(* IEC 61131-3 sources: SortJet_MasterSPS_Aufbau.fbsproj/Device.device.xml.v3^/Plc Logic.plclogic.xml.v3^/Application.application.xml.v3^/09_Station/Stationen/Förderer[202,203]/0_Konfig, 6 files *)

(* ---- Antriebsinformationen_202.gvl ---- *)
(* METADATA
{
	"v3Meta": {
		"objectGuid": "ae52444f-d7c0-4b01-95e4-d9e00420f7a3"
	}
}
*)
{attribute 'allow_unqualified_access'}
NAMESPACE Antriebsinformationen_202
VAR_GLOBAL

//**************************************************************************************************)
// ANTRIEBSINFORMATION  *)
//**************************************************************************************************)

  apgInfoStation202Glastransport : ARRAY[cWAND_1..cANZAHL_WAENDE] OF AntriebsInformationen := [
    (
      wAchsID                                 :=      12,  // Achs ID aus dem EConSet
      stTyp                                   := 'Belt',  // Typ
      wpSchaltschrank                         :=   2020,  // Daten aus dem Schaltplan
      wpSchaltplanreihe                       :=      2,  // Daten aus dem Schaltplan
      wpSchaltplanseite                       :=    100,  // Daten aus dem Schaltplan
      rpMaxGeschwindigkeit                    :=   1000,  // [mm/s]   Max- Geschwindigkeit für den Automatikbetrieb
      rpHandGeschwindigkeit                   :=    333,  // [mm/s]   Hand- Geschwindigkeit
      rpReduzierteGeschwindigkeit             :=    250,  // [mm/s]   Reduzierte Geschwindigkeit
      rpReferenzGeschwindigkeit               :=    100,  // [mm/s]   Geschwindigkeit für die Referenzfahrt
      rpEinrichtGeschwindigkeit               :=     50,  // [mm/s]   Max Geschwindigkeit während der Einrichtung der Anlage
      rpMaxBeschleunigung                     :=   1500,  // [mm/s^2] Max Beschleunigung
      rpMaxVerzoegerung                       :=   2000,  // [mm/s^2] Max Verzoegerung
      rpMaxRuckzeit                           :=     50,  // [ms]     Ruckzeit des Antriebs
      rpReduzierteBeschleunigung              :=   1000,  // [mm/s^2] Reduzierte Beschleunigung
      rpReduzierteVerzoegerung                :=   1000,  // [mm/s^2] Reduzierte Verzoegerung
      rpBeschleunigungFremdanlage             :=   1000,  // [mm/s^2] Beschleunigung zu einer Fremdanlage
      rpGeschwindigkeitMessen                 :=    667,  // [mm/s] Geschwindigkeit beim Scheiben messen
      rpGeschwindigkeitSystemcheck            :=  500.0,  // [mm/s]   Geschwindigkeit im Systemcheck (nur Glastransport)
      rpGeschwindigkeitSystemcheckReduzierung :=  167.0,  // [mm/s]   Geschwindigkeit im Systemcheck bei belegtem Vorstop-Sensor (nur Glastransport)
      stOptionen                              := ( eEndschalterQuelle    := Endschalterquelle_EN.KEINE,     // Hardware-Endschalter: KEINE, UMRICHTER oder SPS
                                                   bVersorgungUeberXVR   := FALSE,                          // XVR-Modus: brueckt Hauptschalter 400 V und LS 230 V
                                                   bBremseLoesenFreigabe := FALSE )                         // Der Antrieb darf über eine Betriebsart die Bremse lösen
    )];

  apgInfoStation202Glastransport_Slave : ARRAY[cWAND_1..cANZAHL_WAENDE] OF AntriebsInformationen := [
    (
      wAchsID                                 :=     65,  // Achs ID aus dem EConSet
      stTyp                                   := 'Belt',  // Typ
      wpSchaltschrank                         :=   2021,  // Daten aus dem Schaltplan
      wpSchaltplanreihe                       :=     02,  // Daten aus dem Schaltplan
      wpSchaltplanseite                       :=    100,  // Daten aus dem Schaltplan
      rpMaxGeschwindigkeit                    :=      0,  // [mm/s]   Max- Geschwindigkeit für den Automatikbetrieb
      rpHandGeschwindigkeit                   :=      0,  // [mm/s]   Hand- Geschwindigkeit
      rpReduzierteGeschwindigkeit             :=      0,  // [mm/s]   Reduzierte Geschwindigkeit
      rpReferenzGeschwindigkeit               :=      0,  // [mm/s]   Geschwindigkeit für die Referenzfahrt
      rpEinrichtGeschwindigkeit               :=      0,  // [mm/s]   Max Geschwindigkeit während der Einrichtung der Anlage
      rpMaxBeschleunigung                     :=      0,  // [mm/s^2] Max Beschleunigung
      rpMaxVerzoegerung                       :=      0,  // [mm/s^2] Max Verzoegerung
      rpMaxRuckzeit                           :=      0,  // [ms]     Ruckzeit des Antriebs
      rpReduzierteBeschleunigung              :=      0,  // [mm/s^2] Reduzierte Beschleunigung
      rpReduzierteVerzoegerung                :=      0,  // [mm/s^2] Reduzierte Verzoegerung
      rpBeschleunigungFremdanlage             :=      0,  // [mm/s^2] Beschleunigung zu einer Fremdanlage
      rpGeschwindigkeitMessen                 :=      0,  // [mm/s] Geschwindigkeit beim Scheiben messen
      rpGeschwindigkeitSystemcheck            :=  500.0,  // [mm/s]   Geschwindigkeit im Systemcheck (nur Glastransport)
      rpGeschwindigkeitSystemcheckReduzierung :=  167.0,  // [mm/s]   Geschwindigkeit im Systemcheck bei belegtem Vorstop-Sensor (nur Glastransport)
      stOptionen                              := ( eEndschalterQuelle    := Endschalterquelle_EN.KEINE,     // Hardware-Endschalter: KEINE, UMRICHTER oder SPS
                                                   bVersorgungUeberXVR   := FALSE,                          // XVR-Modus: brueckt Hauptschalter 400 V und LS 230 V
                                                   bBremseLoesenFreigabe := FALSE )                         // Der Antrieb darf über eine Betriebsart die Bremse lösen
    )];

  apgInfoStation202Kippen : AntriebsInformationen :=
    (
      wAchsID                                 :=     65,  // Achs ID aus dem EConSet
      stTyp                                   := 'Tilt',  // Typ
      wpSchaltschrank                         :=      0,  // Daten aus dem Schaltplan
      wpSchaltplanreihe                       :=     02,  // Daten aus dem Schaltplan
      wpSchaltplanseite                       :=      0,  // Daten aus dem Schaltplan
      rpMaxGeschwindigkeit                    :=      0,  // [Grad/s]   Max- Geschwindigkeit für den Automatikbetrieb
      rpHandGeschwindigkeit                   :=      0,  // [Grad/s]   Hand- Geschwindigkeit
      rpReduzierteGeschwindigkeit             :=      0,  // [Grad/s]   Reduzierte Geschwindigkeit
      rpReferenzGeschwindigkeit               :=      0,  // [Grad/s]   Geschwindigkeit für die Referenzfahrt
      rpEinrichtGeschwindigkeit               :=      0,  // [Grad/s]   Max Geschwindigkeit während der Einrichtung der Anlage
      rpMaxBeschleunigung                     :=      0,  // [Grad/s^2] Max Beschleunigung
      rpMaxVerzoegerung                       :=      0,  // [Grad/s^2] Max Verzoegerung
      rpMaxRuckzeit                           :=      0,  // [ms] Ruckzeit des Antriebs
      rpReduzierteBeschleunigung              :=      0,  // [Grad/s^2] Reduzierte Beschleunigung
      rpReduzierteVerzoegerung                :=      0,  // [Grad/s^2] Reduzierte Verzoegerung
      rpBeschleunigungFremdanlage             :=      0,  // [Grad/s^2] Beschleunigung zu einer Fremdanlage
      rpGeschwindigkeitMessen                 :=      0,  // [Grad/s] Geschwindigkeit beim Scheiben messen
      rpGeschwindigkeitSystemcheck            :=  500.0,  // [mm/s]   Geschwindigkeit im Systemcheck (nur Glastransport)
      rpGeschwindigkeitSystemcheckReduzierung :=  167.0,  // [mm/s]   Geschwindigkeit im Systemcheck bei belegtem Vorstop-Sensor (nur Glastransport)
      stOptionen                              := ( eEndschalterQuelle    := Endschalterquelle_EN.KEINE,     // Hardware-Endschalter: KEINE, UMRICHTER oder SPS
                                                   bVersorgungUeberXVR   := FALSE,                          // XVR-Modus: brueckt Hauptschalter 400 V und LS 230 V
                                                   bBremseLoesenFreigabe := FALSE )                         // Der Antrieb darf über eine Betriebsart die Bremse lösen
    );

  // Querfahrt
  apgInfoStation202Querfahrt : AntriebsInformationen :=
    (
      wAchsID                                 :=        65,  // Achs ID aus dem EConSet
      stTyp                                   := 'Lateral',  // Typ
      wpSchaltschrank                         :=      2113,  // Daten aus dem Schaltplan
      wpSchaltplanreihe                       :=        02,  // Daten aus dem Schaltplan
      wpSchaltplanseite                       :=         0,  // Daten aus dem Schaltplan
      rpMaxGeschwindigkeit                    :=      1000,  // [mm/s]   Max- Geschwindigkeit für den Automatikbetrieb
      rpHandGeschwindigkeit                   :=      1000,  // [mm/s]   Hand- Geschwindigkeit
      rpReduzierteGeschwindigkeit             :=        25,  // [mm/s]   Reduzierte Geschwindigkeit
      rpReferenzGeschwindigkeit               :=        10,  // [mm/s]   Geschwindigkeit für die Referenzfahrt
      rpEinrichtGeschwindigkeit               :=        10,  // [mm/s]   Max Geschwindigkeit während der Einrichtung der Anlage
      rpMaxBeschleunigung                     :=       500,  // [mm/s^2] Max Beschleunigung
      rpMaxVerzoegerung                       :=       500,  // [mm/s^2] Max Verzoegerung
      rpMaxRuckzeit                           :=      1000,  // [ms]     Ruckzeit des Antriebs
      rpReduzierteBeschleunigung              :=        10,  // [mm/s^2] Reduzierte Beschleunigung
      rpReduzierteVerzoegerung                :=        10,  // [mm/s^2] Reduzierte Verzoegerung
      rpBeschleunigungFremdanlage             :=         0,  // [mm/s^2] Beschleunigung zu einer Fremdanlage
      rpGeschwindigkeitMessen                 :=         0,  // [mm/s] Geschwindigkeit beim Scheiben messen
      rpGeschwindigkeitSystemcheck            :=     500.0,  // [mm/s]   Geschwindigkeit im Systemcheck (nur Glastransport)
      rpGeschwindigkeitSystemcheckReduzierung :=     167.0,  // [mm/s]   Geschwindigkeit im Systemcheck bei belegtem Vorstop-Sensor (nur Glastransport)
      stOptionen                              := ( eEndschalterQuelle    := Endschalterquelle_EN.UMRICHTER, // Hardware-Endschalter: KEINE, UMRICHTER oder SPS
                                                   bVersorgungUeberXVR   := FALSE,                          // XVR-Modus: brueckt Hauptschalter 400 V und LS 230 V
                                                   bBremseLoesenFreigabe := FALSE )                         // Der Antrieb darf über eine Betriebsart die Bremse lösen
    );

END_VAR

END_NAMESPACE

(* ---- Antriebsinformationen_203.gvl ---- *)
(* METADATA
{
	"v3Meta": {
		"objectGuid": "bcc74c11-83af-44f4-ba61-cf23f0f94a5f"
	}
}
*)
{attribute 'allow_unqualified_access'}
NAMESPACE Antriebsinformationen_203
VAR_GLOBAL

//**************************************************************************************************)
// ANTRIEBSINFORMATION  *)
//**************************************************************************************************)

  apgInfoStation203Glastransport : ARRAY[cWAND_1..cANZAHL_WAENDE] OF AntriebsInformationen := [
    (
      wAchsID                                 :=     11,   // Achs ID aus dem EConSet
      stTyp                                   := 'Belt',  // Typ
      wpSchaltschrank                         :=   2030,  // Daten aus dem Schaltplan
      wpSchaltplanreihe                       :=      2,  // Daten aus dem Schaltplan
      wpSchaltplanseite                       :=    100,  // Daten aus dem Schaltplan
      rpMaxGeschwindigkeit                    :=   1000,  // [mm/s]   Max- Geschwindigkeit für den Automatikbetrieb
      rpHandGeschwindigkeit                   :=    333,  // [mm/s]   Hand- Geschwindigkeit
      rpReduzierteGeschwindigkeit             :=     67,  // [mm/s]   Reduzierte Geschwindigkeit
      rpReferenzGeschwindigkeit               :=      0,  // [mm/s]   Geschwindigkeit für die Referenzfahrt
      rpEinrichtGeschwindigkeit               :=     50,  // [mm/s]   Max Geschwindigkeit während der Einrichtung der Anlage
      rpMaxBeschleunigung                     :=   1500,  // [mm/s^2] Max Beschleunigung
      rpMaxVerzoegerung                       :=   2000,  // [mm/s^2] Max Verzoegerung
      rpMaxRuckzeit                           :=     50,  // [ms]     Ruckzeit des Antriebs
      rpReduzierteBeschleunigung              :=   1000,  // [mm/s^2] Reduzierte Beschleunigung
      rpReduzierteVerzoegerung                :=   1000,  // [mm/s^2] Reduzierte Verzoegerung
      rpBeschleunigungFremdanlage             :=   1000,  // [mm/s^2] Beschleunigung zu einer Fremdanlage
      rpGeschwindigkeitMessen                 :=    667,  // [mm/s] Geschwindigkeit beim Scheiben messen
      rpGeschwindigkeitSystemcheck            :=  500.0,  // [mm/s]   Geschwindigkeit im Systemcheck (nur Glastransport)
      rpGeschwindigkeitSystemcheckReduzierung :=  167.0,  // [mm/s]   Geschwindigkeit im Systemcheck bei belegtem Vorstop-Sensor (nur Glastransport)
      stOptionen                              := ( eEndschalterQuelle    := Endschalterquelle_EN.KEINE,     // Hardware-Endschalter: KEINE, UMRICHTER oder SPS
                                                   bVersorgungUeberXVR   := FALSE,                          // XVR-Modus: brueckt Hauptschalter 400 V und LS 230 V
                                                   bBremseLoesenFreigabe := FALSE )                         // Der Antrieb darf über eine Betriebsart die Bremse lösen
    )];

  apgInfoStation203Glastransport_Slave : ARRAY[cWAND_1..cANZAHL_WAENDE] OF AntriebsInformationen := [
    (
      wAchsID                                 :=     65,  // Achs ID aus dem EConSet
      stTyp                                   := 'Belt',  // Typ
      wpSchaltschrank                         :=   2031,  // Daten aus dem Schaltplan
      wpSchaltplanreihe                       :=     02,  // Daten aus dem Schaltplan
      wpSchaltplanseite                       :=    100,  // Daten aus dem Schaltplan
      rpMaxGeschwindigkeit                    :=      0,  // [mm/s]   Max- Geschwindigkeit für den Automatikbetrieb
      rpHandGeschwindigkeit                   :=      0,  // [mm/s]   Hand- Geschwindigkeit
      rpReduzierteGeschwindigkeit             :=      0,  // [mm/s]   Reduzierte Geschwindigkeit
      rpReferenzGeschwindigkeit               :=      0,  // [mm/s]   Geschwindigkeit für die Referenzfahrt
      rpEinrichtGeschwindigkeit               :=      0,  // [mm/s]   Max Geschwindigkeit während der Einrichtung der Anlage
      rpMaxBeschleunigung                     :=      0,  // [mm/s^2] Max Beschleunigung
      rpMaxVerzoegerung                       :=      0,  // [mm/s^2] Max Verzoegerung
      rpMaxRuckzeit                           :=      0,  // [ms]     Ruckzeit des Antriebs
      rpReduzierteBeschleunigung              :=      0,  // [mm/s^2] Reduzierte Beschleunigung
      rpReduzierteVerzoegerung                :=      0,  // [mm/s^2] Reduzierte Verzoegerung
      rpBeschleunigungFremdanlage             :=      0,  // [mm/s^2] Beschleunigung zu einer Fremdanlage
      rpGeschwindigkeitMessen                 :=      0,  // [mm/s] Geschwindigkeit beim Scheiben messen
      rpGeschwindigkeitSystemcheck            :=  500.0,  // [mm/s]   Geschwindigkeit im Systemcheck (nur Glastransport)
      rpGeschwindigkeitSystemcheckReduzierung :=  167.0,  // [mm/s]   Geschwindigkeit im Systemcheck bei belegtem Vorstop-Sensor (nur Glastransport)
      stOptionen                              := ( eEndschalterQuelle    := Endschalterquelle_EN.KEINE,     // Hardware-Endschalter: KEINE, UMRICHTER oder SPS
                                                   bVersorgungUeberXVR   := FALSE,                          // XVR-Modus: brueckt Hauptschalter 400 V und LS 230 V
                                                   bBremseLoesenFreigabe := FALSE )                         // Der Antrieb darf über eine Betriebsart die Bremse lösen
    )];

  apgInfoStation203Kippen : AntriebsInformationen :=
    (
      wAchsID                                 :=     65,  // Achs ID aus dem EConSet
      stTyp                                   := 'Tilt',  // Typ
      wpSchaltschrank                         :=      0,  // Daten aus dem Schaltplan
      wpSchaltplanreihe                       :=     02,  // Daten aus dem Schaltplan
      wpSchaltplanseite                       :=      0,  // Daten aus dem Schaltplan
      rpMaxGeschwindigkeit                    :=      0,  // [Grad/s]   Max- Geschwindigkeit für den Automatikbetrieb
      rpHandGeschwindigkeit                   :=      0,  // [Grad/s]   Hand- Geschwindigkeit
      rpReduzierteGeschwindigkeit             :=      0,  // [Grad/s]   Reduzierte Geschwindigkeit
      rpReferenzGeschwindigkeit               :=      0,  // [Grad/s]   Geschwindigkeit für die Referenzfahrt
      rpEinrichtGeschwindigkeit               :=      0,  // [Grad/s]   Max Geschwindigkeit während der Einrichtung der Anlage
      rpMaxBeschleunigung                     :=      0,  // [Grad/s^2] Max Beschleunigung
      rpMaxVerzoegerung                       :=      0,  // [Grad/s^2] Max Verzoegerung
      rpMaxRuckzeit                           :=      0,  // [ms] Ruckzeit des Antriebs
      rpReduzierteBeschleunigung              :=      0,  // [Grad/s^2] Reduzierte Beschleunigung
      rpReduzierteVerzoegerung                :=      0,  // [Grad/s^2] Reduzierte Verzoegerung
      rpBeschleunigungFremdanlage             :=      0,  // [Grad/s^2] Beschleunigung zu einer Fremdanlage
      rpGeschwindigkeitMessen                 :=      0,  // [Grad/s] Geschwindigkeit beim Scheiben messen
      rpGeschwindigkeitSystemcheck            :=  500.0,  // [mm/s]   Geschwindigkeit im Systemcheck (nur Glastransport)
      rpGeschwindigkeitSystemcheckReduzierung :=  167.0,  // [mm/s]   Geschwindigkeit im Systemcheck bei belegtem Vorstop-Sensor (nur Glastransport)
      stOptionen                              := ( eEndschalterQuelle    := Endschalterquelle_EN.KEINE,     // Hardware-Endschalter: KEINE, UMRICHTER oder SPS
                                                   bVersorgungUeberXVR   := FALSE,                          // XVR-Modus: brueckt Hauptschalter 400 V und LS 230 V
                                                   bBremseLoesenFreigabe := FALSE )                         // Der Antrieb darf über eine Betriebsart die Bremse lösen
    );

  // Querfahrt
  apgInfoStation203Querfahrt : AntriebsInformationen :=
    (
      wAchsID                                 :=        65,  // Achs ID aus dem EConSet
      stTyp                                   := 'Lateral',  // Typ
      wpSchaltschrank                         :=      2113,  // Daten aus dem Schaltplan
      wpSchaltplanreihe                       :=        02,  // Daten aus dem Schaltplan
      wpSchaltplanseite                       :=         0,  // Daten aus dem Schaltplan
      rpMaxGeschwindigkeit                    :=      1000,  // [mm/s]   Max- Geschwindigkeit für den Automatikbetrieb
      rpHandGeschwindigkeit                   :=      1000,  // [mm/s]   Hand- Geschwindigkeit
      rpReduzierteGeschwindigkeit             :=        25,  // [mm/s]   Reduzierte Geschwindigkeit
      rpReferenzGeschwindigkeit               :=        10,  // [mm/s]   Geschwindigkeit für die Referenzfahrt
      rpEinrichtGeschwindigkeit               :=        10,  // [mm/s]   Max Geschwindigkeit während der Einrichtung der Anlage
      rpMaxBeschleunigung                     :=       500,  // [mm/s^2] Max Beschleunigung
      rpMaxVerzoegerung                       :=       500,  // [mm/s^2] Max Verzoegerung
      rpMaxRuckzeit                           :=      1000,  // [ms]     Ruckzeit des Antriebs
      rpReduzierteBeschleunigung              :=        10,  // [mm/s^2] Reduzierte Beschleunigung
      rpReduzierteVerzoegerung                :=        10,  // [mm/s^2] Reduzierte Verzoegerung
      rpBeschleunigungFremdanlage             :=         0,  // [mm/s^2] Beschleunigung zu einer Fremdanlage
      rpGeschwindigkeitMessen                 :=         0,  // [mm/s] Geschwindigkeit beim Scheiben messen
      rpGeschwindigkeitSystemcheck            :=     500.0,  // [mm/s]   Geschwindigkeit im Systemcheck (nur Glastransport)
      rpGeschwindigkeitSystemcheckReduzierung :=     167.0,  // [mm/s]   Geschwindigkeit im Systemcheck bei belegtem Vorstop-Sensor (nur Glastransport)
      stOptionen                              := ( eEndschalterQuelle    := Endschalterquelle_EN.UMRICHTER, // Hardware-Endschalter: KEINE, UMRICHTER oder SPS
                                                   bVersorgungUeberXVR   := FALSE,                          // XVR-Modus: brueckt Hauptschalter 400 V und LS 230 V
                                                   bBremseLoesenFreigabe := FALSE )                         // Der Antrieb darf über eine Betriebsart die Bremse lösen
    );

END_VAR

END_NAMESPACE

(* ---- MK_Station_202.gvl ---- *)
(* METADATA
{
	"v3Meta": {
		"objectGuid": "7b2503c5-79dd-46b3-9fd2-96547eeb48a2"
	}
}
*)
{attribute 'allow_unqualified_access'}
NAMESPACE MK_Station_202
VAR_GLOBAL

//-------------------------------------------------------------------------------------------------
// MASCHINEPARAMETER: SENKRECHTFOERDERER
//-------------------------------------------------------------------------------------------------

  apgMKStation202 : Parameter_Station:=
    (
      stStationsNummern                     := ( NummerIntern :=   202,                                                      // Stationsnummer fuer das MMI und die Stationsangabe der Meldungen
                                                 NummerExtern :=  1202,                                                      // Stationsnummer fuer Bedienermeldungen
                                                 NummerSPS    :=   202 ),                                                    // Stationsnummer SPS-intern (Indizes)
      bDeaktivieren                         := FALSE,                                                                        // Station deaktiviert (keine Auftraege, keine Referenzfahrt)
      wMeldungsNummer                       := 1720,                                                                         // Basis-Meldungsnummer (WatchIO)
      eStationsTyp                          := eStation,                                                                     // Typ der Station
      eaAutomatikkreis                      := [eAutomatikkreis_1],                                                          // Automatikkreise, zu denen die Station gehoert
      eaSicherheitskreis                    := [eSicherheitskreis_Undefiniert],                                              // Sicherheitskreise, in die die Station eingebunden ist
      // astSicherheitskreisTeilabschaltung
      eSystemcheckZyklus                    := eSystemcheckZyklus_1,                                                         // In welchem Zyklus des Systemchecks die Station geprueft wird
      stSchnittstellendaten                 := ( wVorgaengerStation := cSTATION_201,                                         // Station vor dieser Station (cSTATION_DYNAMISCH bei mehreren)
                                                 wNachfolgerStation := cSTATION_203,                                         // Station nach dieser Station (cSTATION_DYNAMISCH bei mehreren)
                                                 bStationIstShuttle := FALSE                                                 // Station ist ein Shuttle
                                               ),
      stStationsOptionen                    := ( stSystemcheck :=  ( bScheibenVermessenSystemCheck               := TRUE,    // Scheiben im Systemcheck vermessen
                                                                     bScheibeNachSystemcheckAufAuslauf           := TRUE,    // Scheibe nach dem Systemcheck auf den Auslaufsensor fahren
                                                                     bSystemCheckMitVorgaengerBatchTransport     := FALSE,   // derzeit ohne Funktion
                                                                     bSystemCheckMitNachfolgerBatchTransport     := FALSE,   // derzeit ohne Funktion
                                                                     bOptionSystemCheckScheibeMittigLegen        := FALSE ), // derzeit ohne Funktion

                                                 // stTransfershuttle
                                                 stGlastransport :=  ( bVortransport                             := FALSE,   // Vortransport aktivieren [Bsp.: Nach einem Eintransport mit gesetztem Bit <Letzte Scheibe>]
                                                                       bTransportMasterSlaveEintransport         := FALSE,   // derzeit ohne Funktion
                                                                       bTransportMasterSlaveAustransport         := TRUE ,   // Austransport als Slave auf die Achse des Nachfolgers
                                                                       bGLasUebernahmeSenkrecht                  := FALSE,   // RKT - Eintransport in Senkrechter-Position bzw. in Waagerechter- Position [default]
                                                                       bAustransportISOLinie                     := FALSE,   // Austransport an eine ISO-Linie
                                                                       bScheibenVermessen                        := FALSE,   // Scheibenmessung am Anlegetisch/Anlegewand
                                                                       bMessrichtungNegativ                      := FALSE,   // Negative Fahrtrichtung beim Messen
                                                                       bScheibenmessungEintransport              := FALSE,   // Scheibenmessung beim Eintransport
                                                                       bScheibenmessungSensorVorabAuslauf        := FALSE    // Scheibenmessung mit SensorVorabAuslauf z.B. Anlegewand
                                                                      ),
                                                 // stAnlegetisch
                                                 // stEckuebergabe
                                                 // stDrehstation
                                                 bVorAbKomponentenAnsteuerung              := FALSE,                         // VorAbKomponentenAnsteuerung Auftraege werden bearbeitet
                                                 bVerstellungEinAusGefahrenLogikDrehen     := FALSE,                         // Verstellung: Logik ein-/ausgefahren gedreht
                                                 bLangsamfahrtNockenQuerfahrtAktivieren    := FALSE,                         // Querfahrt: Langsamfahrt-Nocken auswerten
                                                 bSKBlockierenDurchVorabSensoren           := FALSE,                         // Vorab-Sensoren belegt blockieren das Oeffnen des Sicherheitskreises
                                                 bStationLeerfahrenBeiSkAnforderung        := FALSE,                         // Station bei Anforderung Sicherheitskreis leerfahren
                                                 bGlasAbgenommenAutomatischQuittieren      := FALSE,                         // derzeit ohne Funktion
                                                 bScheibeAbnehmenNachEintransport          := FALSE                          // Scheibe nach dem Eintransport wieder abnehmen
                                               ),
      stStationsAufbau                      := ( bGeblase                      := [ cANZAHL_WAENDE(FALSE) ],                 // Ausbaustufe: Geblaese je Wand
                                                 bGlastransport                := [ TRUE ],                                  // Ausbaustufe: Glastransport je Wand
                                                 bKippen                       := [ cANZAHL_WAENDE(FALSE) ],                 // Ausbaustufe: Kippen je Wand
                                                 bKippenSchuetz                := FALSE,                                     // Kippen ueber Schuetz statt Umrichter
                                                 bTransportVerstellung         := [ cANZAHL_WAENDE(FALSE) ],                 // Ausbaustufe Shuttle: Transport-/Dickenverstellung je Wand
                                                 bHub                          := FALSE,                                     // Ausbaustufe: Hub der Station
                                                 bHubrahmen                    := FALSE,                                     // Ausbaustufe: Hubrahmen (Riemen heben/senken)
                                                 bDrehen                       := FALSE,                                     // Ausbaustufe: Drehen
                                                 bQuerachse                    := FALSE,                                     // Ausbaustufe: Querachse
                                                 bMessachse                    := FALSE,                                     // Ausbaustufe: Messachse (Anlegetisch, Anlegewand)
                                                 bDruckluft                    := FALSE,                                     // Druckluftueberwachung vorhanden
                                                 bAnschlag                     := FALSE,                                     // Ausbaustufe: Ausrichtanschlaege
                                                 bSensorAuslauf                := TRUE,                                      // Auslaufsensor vorhanden
                                                 bSensorEinlauf                := TRUE,                                      // Einlaufsensor vorhanden
                                                 bSensorEinlaufStopp           := FALSE,                                     // Shuttle: zusaetzlicher Stopp-Sensor am Einlauf (ohne: Einlaufsensor), Gegenstueck zum Auslauf-Stopp im Rueckwaertstransport
                                                 bSensorAuslaufStopp           := FALSE,                                     // Shuttle: zusaetzlicher Stopp-Sensor am Auslauf (ohne: Auslaufsensor), Verfahrfreigabe und Scheibe hat Shuttle verlassen
                                                 bDurchlaufSperreZumNachfolger := FALSE,                                     // Ausbaustufe: bewegliche Abschrankung zum Nachfolger
                                                 bQuerfahrt                    := FALSE,                                     // Ausbaustufe: Querfahrt
                                                 bKipparme                     := FALSE,                                     // Ausbaustufe: Kipparme
                                                 bSlaveAntrieb                 := FALSE,                                     // Glastransport mit Slave-Antrieb
                                                 bMessachseAmEndeVomTisch      := FALSE,                                     // Messachse am Ende des Tisches (Hoehenfehler fragt den Bediener)
                                                 bWandverstellung              := [ FALSE ],                                 // Ausbaustufe Station: Wandverstellung je Wand
                                                 bWandverstellungMotorisch     := FALSE,                                     // Shuttle: Transport-/Wandverstellung mit Antrieb statt pneumatisch
                                                 bRoellchenleiste              := [ FALSE ],                                 // Ausbaustufe Station: Roellchenleiste je Wand
                                                 bDurchgang                    := FALSE,                                     // Station ist Teil eines Durchgangs (belegt = Oeffnen blockiert)
                                                 bRolltor                      := FALSE,                                     // Ausbaustufe Faecherwagen: Rolltor
                                                 bKlemmzylinder                := FALSE,                                     // Ausbaustufe Faecherwagen: Klemmzylinder fixiert den Oberrahmen beim Ein- und Ausschleusen
                                                 bGreifer                      := [cANZAHL_WAENDE(FALSE)],                   // Shuttle: Greifer je Wand (Scheibe aus dem Faecherwagen ziehen bzw. hineinschieben)
                                                 bRFID                         := FALSE,                                     // RFID-Leser vorhanden
                                                 bAGV                          := FALSE,                                     // Ausbaustufe Faecherwagen: Betrieb mit AGV
                                                 bDLSSchmiersystem             := FALSE,                                     // Zentralschmierung DLS vorhanden
                                                 bGlastransportSlaveVorhanden  := FALSE,                                     // Glastransport mit Slave-Antrieb (Meldungen/Ueberwachung Slave)
                                                 wHydraulikstation             := 0                                          // Faecherwagen Hydraulik: zugeordnete Hydraulikstation (cHYDRAULIKSTATION_x), 0 = keine
                                               ),
      stStationsParameter                   := ( rLaengeUebergroesseScheibe              := 3300,                            // Shuttle: ab dieser Scheibenlaenge gilt die Scheibe als uebergross [mm]
                                                 rMinGlasHoeheAutomatischenEintransport  := 500,                             // VSG: Mindesthoehe fuer automatischen Eintransport [mm]
                                                 rMinGlasLaengeAutomatischenEintransport := 500,                             // VSG: Mindestlaenge fuer automatischen Eintransport [mm]
                                                 wMaximaleAnzahlAktiverAuftraege := 1,                                       // derzeit ohne Funktion
                                                 rMinPosSwEsEingrenzung                  := 0.0,                             // Externer zusaetzlicher Software-Endschalter MIN; 0 = inaktiv; darf den MK-MIN nur weiter eingrenzen
                                                 rMaxPosSwEsEingrenzung                  := 0.0,                             // Externer zusaetzlicher Software-Endschalter MAX; 0 = inaktiv; darf den MK-MAX nur weiter eingrenzen
                                                 rPosFreigabePufferAusfahren             := 0.0                              // derzeit ohne Funktion
                                              ),
      // stFremdanlage
      stGlasdaten                           := [( rlMinGlasLaenge := 350,                                                    // minimal zulässige GlasLänge
                                                  rlMaxGlasLaenge := 2500,                                                   // maximale zulässige GlasLänge
                                                  rlMinGlasHoehe  := 190,                                                    // minimal zulässige GlasHöhe
                                                  rlMaxGlasHoehe  := 1800,                                                   // maximale zulässige GlasHöhe
                                                  rlMinGlasDicke  := 3,                                                    // minimal zulässige GlasDicke
                                                  rlMaxGlasDicke  := 12.76,                                                     // maximal zulaessige Glasdicke [mm]
                                                  rlLaengeMaxGlas := 0.0                                                     // maximal zulaessige Glaslaenge [mm]
                                               )]
      // astShuttleAnhaltenQuellen
    );

  apgMKStation202Glastransport : ARRAY[cWAND_1..cANZAHL_WAENDE] OF Parameter_Glastransport := [
    (
      rLaengeStation                        := 4600, // Länge der Station
      rScheibenabstand                      :=  300, // Der Abstand zwischen zwei Scheiben auf der Station
      rWegUeberEinlauf                      :=   50, // Weg ueber den Einlaufsensor hinaus [mm]
      rWegUeberAuslauf                      :=   50, // Weg ueber den Auslaufsensor hinaus [mm]
      rWegUeberSensorenSystemCheck          :=   15, // Der Weg der Ueber ein die Sensoren zum vermessen der Scheiben
      rUeberwachungAuslaufsensor            :=  500, // Ueberwachung des Auslaufsensors [Strecke in der der Auslaufsensor Frei / ueberfahren werden soll]
      rUeberwachungEinlaufsensor            :=  500, // Ueberwachung des Einlaufsensors [Strecke in der der Einlaufsensor Frei / ueberfahren werden soll]
      rWegUeberEinlaufEintransport          :=   80, // Eintransport vorwaerts: Abstand Scheibenhinterkante zum Einlaufsensor [mm]
      rWegUeberEinlaufAustransport          :=   50, // Lage Auf Einlauf: Scheibe liegt um diesen Weg auf dem Einlaufsensor [mm]
      rWegUeberAuslaufEintransport          :=   50, // Eintransport rueckwaerts: Abstand Scheibenhinterkante zum Auslaufsensor [mm]
      rWegUeberAuslaufAustransport          :=   50, // Lage Auf Auslauf: Weg ueber den Auslaufsensor hinaus [mm]
      rWegEinlaufsensorZuVorStopSensor      := 4500, // Beschreibt den Weg vum eine Scheibe beim EIntransport vom Einlaufsensor bis ueberden Vorabstopsensor zu verfahren
      rMesstoleranz                         :=   10, // Toleranz-Mass fuer die Scheibenlaengenmessung
      rMessstrecke                          := 4535, // Beschreibt die Strecke ziwischen 2 Sensoren die der Antrieb verfaehrt
      rWegstreckeBisZurVerzoegerung         := 4000  // Beschreibt die Strecke die gefahren werden soll bis der Antrieb abgebremst werden soll, dies gilt fuer Eintransportauftraege die das Bit "Letzte Scheibe" gesetzt haben
    )];

  apgMKStation202Kippen : ARRAY[cWAND_1..cANZAHL_WAENDE] OF Parameter_Kippen := [
    (
      tZeitlicheUeberwachungKippen          := TIME#5000MS, // [ms \ s] Verwendet fuer Antriebe die Ueber einen Schuetz angesteuert werden
      tZeitAntriebsfreigabeErhalten         := TIME#180S,   // [ms \ s] Energieeinsparrung: Zeiteinheit nach der die Antriebsfreigabe entzogen werden soll wenn keine Aktion ansteht [1 s = 1000 ms ]
      rToleranz                             := 0,           // Toleranz beim Entscheiden der aktuellen Position
      rPosition0Grad                        := 0,           // Waagerechte- Position 0 Grad: Position auf die die Station gehoben werden soll
      rPosition84Grad                       := 0,           // Senkrechte- Position 84 Grad: Position auf die die Station gehoben werden soll
      rPosition90Grad                       := 0,           // Senkrechte-Position 90 Grad : Position auf die die Station gesenkt werden soll
      rPosition96Grad                       := 0,           // Senkrechte-Position 96 Grad : Position auf die die Station gesenkt werden soll
      bKippenMitSchuetz                     := TRUE,        // Kippen per Umrichter oder Schütz
      rPosition88_5Grad                     := 0.0          // Senkrechte- Position 84 Grad: Position auf die die Station gehoben werden soll
    )];

   apgMKStation202Querfahrt : Parameter_Querfahrt :=
    (
      tZeitAntriebsfreigabeErhalten          := T#3M // Energieeinsparung: Zeit nach der die Antriebsfreigabe entzogen wird, wenn keine Aktion ansteht
    );

END_VAR
END_NAMESPACE

(* ---- MK_Station_203.gvl ---- *)
(* METADATA
{
	"v3Meta": {
		"objectGuid": "c357eb5d-995e-48ac-a8b0-c12f67a0f286"
	}
}
*)
{attribute 'allow_unqualified_access'}
NAMESPACE MK_Station_203
VAR_GLOBAL

//-------------------------------------------------------------------------------------------------
// MASCHINEPARAMETER: SENKRECHTFOERDERER
//-------------------------------------------------------------------------------------------------

  apgMKStation203 : Parameter_Station:=
    (
      stStationsNummern                     := ( NummerIntern :=   203,                                                      // Stationsnummer fuer das MMI und die Stationsangabe der Meldungen
                                                 NummerExtern :=  1203,                                                      // Stationsnummer fuer Bedienermeldungen
                                                 NummerSPS    :=   203 ),                                                    // Stationsnummer SPS-intern (Indizes)
      bDeaktivieren                         := FALSE,                                                                        // Station deaktiviert (keine Auftraege, keine Referenzfahrt)
      wMeldungsNummer                       := 1740,                                                                         // Basis-Meldungsnummer (WatchIO)
      eStationsTyp                          := eStation,                                                                     // Typ der Station
      eaAutomatikkreis                      := [eAutomatikkreis_1],                                                          // Automatikkreise, zu denen die Station gehoert
      eaSicherheitskreis                    := [eSicherheitskreis_3],                                                        // Sicherheitskreise, in die die Station eingebunden ist
      // astSicherheitskreisTeilabschaltung
      eSystemcheckZyklus                    := eSystemcheckZyklus_1,                                                         // In welchem Zyklus des Systemchecks die Station geprueft wird
      stSchnittstellendaten                 := ( wVorgaengerStation := cSTATION_202,                                         // Station vor dieser Station (cSTATION_DYNAMISCH bei mehreren)
                                                 wNachfolgerStation := cSTATION_204,                                         // Station nach dieser Station (cSTATION_DYNAMISCH bei mehreren)
                                                 bStationIstShuttle := FALSE                                                 // Station ist ein Shuttle
                                               ),
      stStationsOptionen                    := ( stSystemcheck :=  ( bScheibenVermessenSystemCheck               := TRUE,    // Scheiben im Systemcheck vermessen
                                                                     bScheibeNachSystemcheckAufAuslauf           := TRUE,    // Scheibe nach dem Systemcheck auf den Auslaufsensor fahren
                                                                     bSystemCheckMitVorgaengerBatchTransport     := FALSE,   // derzeit ohne Funktion
                                                                     bSystemCheckMitNachfolgerBatchTransport     := FALSE,   // derzeit ohne Funktion
                                                                     bOptionSystemCheckScheibeMittigLegen        := FALSE ), // derzeit ohne Funktion

                                                 // stTransfershuttle
                                                 stGlastransport :=  ( bVortransport                             := FALSE,   // Vortransport aktivieren [Bsp.: Nach einem Eintransport mit gesetztem Bit <Letzte Scheibe>]
                                                                       bTransportMasterSlaveEintransport         := FALSE,   // derzeit ohne Funktion
                                                                       bTransportMasterSlaveAustransport         := TRUE ,   // Austransport als Slave auf die Achse des Nachfolgers
                                                                       bGLasUebernahmeSenkrecht                  := FALSE,   // RKT - Eintransport in Senkrechter-Position bzw. in Waagerechter- Position [default]
                                                                       bAustransportISOLinie                     := FALSE,   // Austransport an eine ISO-Linie
                                                                       bScheibenVermessen                        := FALSE,   // Scheibenmessung am Anlegetisch/Anlegewand
                                                                       bMessrichtungNegativ                      := FALSE,   // Negative Fahrtrichtung beim Messen
                                                                       bScheibenmessungEintransport              := FALSE,   // Scheibenmessung beim Eintransport
                                                                       bScheibenmessungSensorVorabAuslauf        := FALSE    // Scheibenmessung mit SensorVorabAuslauf z.B. Anlegewand
                                                                      ),
                                                 // stAnlegetisch
                                                 // stEckuebergabe
                                                 // stDrehstation
                                                 bVorAbKomponentenAnsteuerung              := FALSE,                         // VorAbKomponentenAnsteuerung Auftraege werden bearbeitet
                                                 bVerstellungEinAusGefahrenLogikDrehen     := FALSE,                         // Verstellung: Logik ein-/ausgefahren gedreht
                                                 bLangsamfahrtNockenQuerfahrtAktivieren    := FALSE,                         // Querfahrt: Langsamfahrt-Nocken auswerten
                                                 bSKBlockierenDurchVorabSensoren           := TRUE,                          // Vorab-Sensoren belegt blockieren das Oeffnen des Sicherheitskreises
                                                 bStationLeerfahrenBeiSkAnforderung        := TRUE,                          // Station bei Anforderung Sicherheitskreis leerfahren
                                                 bGlasAbgenommenAutomatischQuittieren      := FALSE,                         // derzeit ohne Funktion
                                                 bScheibeAbnehmenNachEintransport          := FALSE                          // Scheibe nach dem Eintransport wieder abnehmen
                                               ),
      stStationsAufbau                      := ( bGeblase                      := [ cANZAHL_WAENDE(FALSE) ],                 // Ausbaustufe: Geblaese je Wand
                                                 bGlastransport                := [ TRUE ],                                  // Ausbaustufe: Glastransport je Wand
                                                 bKippen                       := [ cANZAHL_WAENDE(FALSE) ],                 // Ausbaustufe: Kippen je Wand
                                                 bKippenSchuetz                := FALSE,                                     // Kippen ueber Schuetz statt Umrichter
                                                 bTransportVerstellung         := [ cANZAHL_WAENDE(FALSE) ],                 // Ausbaustufe Shuttle: Transport-/Dickenverstellung je Wand
                                                 bHub                          := FALSE,                                     // Ausbaustufe: Hub der Station
                                                 bHubrahmen                    := FALSE,                                     // Ausbaustufe: Hubrahmen (Riemen heben/senken)
                                                 bDrehen                       := FALSE,                                     // Ausbaustufe: Drehen
                                                 bQuerachse                    := FALSE,                                     // Ausbaustufe: Querachse
                                                 bMessachse                    := FALSE,                                     // Ausbaustufe: Messachse (Anlegetisch, Anlegewand)
                                                 bDruckluft                    := FALSE,                                     // Druckluftueberwachung vorhanden
                                                 bAnschlag                     := FALSE,                                     // Ausbaustufe: Ausrichtanschlaege
                                                 bSensorAuslauf                := TRUE,                                      // Auslaufsensor vorhanden
                                                 bSensorEinlauf                := TRUE,                                      // Einlaufsensor vorhanden
                                                 bSensorEinlaufStopp           := FALSE,                                     // Shuttle: zusaetzlicher Stopp-Sensor am Einlauf (ohne: Einlaufsensor), Gegenstueck zum Auslauf-Stopp im Rueckwaertstransport
                                                 bSensorAuslaufStopp           := FALSE,                                     // Shuttle: zusaetzlicher Stopp-Sensor am Auslauf (ohne: Auslaufsensor), Verfahrfreigabe und Scheibe hat Shuttle verlassen
                                                 bDurchlaufSperreZumNachfolger := FALSE,                                     // Ausbaustufe: bewegliche Abschrankung zum Nachfolger
                                                 bQuerfahrt                    := FALSE,                                     // Ausbaustufe: Querfahrt
                                                 bKipparme                     := FALSE,                                     // Ausbaustufe: Kipparme
                                                 bSlaveAntrieb                 := FALSE,                                     // Glastransport mit Slave-Antrieb
                                                 bMessachseAmEndeVomTisch      := FALSE,                                     // Messachse am Ende des Tisches (Hoehenfehler fragt den Bediener)
                                                 bWandverstellung              := [ FALSE ],                                 // Ausbaustufe Station: Wandverstellung je Wand
                                                 bWandverstellungMotorisch     := FALSE,                                     // Shuttle: Transport-/Wandverstellung mit Antrieb statt pneumatisch
                                                 bRoellchenleiste              := [ FALSE ],                                 // Ausbaustufe Station: Roellchenleiste je Wand
                                                 bDurchgang                    := TRUE,                                      // Station ist Teil eines Durchgangs (belegt = Oeffnen blockiert)
                                                 bRolltor                      := FALSE,                                     // Ausbaustufe Faecherwagen: Rolltor
                                                 bKlemmzylinder                := FALSE,                                     // Ausbaustufe Faecherwagen: Klemmzylinder fixiert den Oberrahmen beim Ein- und Ausschleusen
                                                 bGreifer                      := [cANZAHL_WAENDE(FALSE)],                   // Shuttle: Greifer je Wand (Scheibe aus dem Faecherwagen ziehen bzw. hineinschieben)
                                                 bRFID                         := FALSE,                                     // RFID-Leser vorhanden
                                                 bAGV                          := FALSE,                                     // Ausbaustufe Faecherwagen: Betrieb mit AGV
                                                 bDLSSchmiersystem             := FALSE,                                     // Zentralschmierung DLS vorhanden
                                                 bGlastransportSlaveVorhanden  := FALSE,                                     // Glastransport mit Slave-Antrieb (Meldungen/Ueberwachung Slave)
                                                 wHydraulikstation             := 0                                          // Faecherwagen Hydraulik: zugeordnete Hydraulikstation (cHYDRAULIKSTATION_x), 0 = keine
                                               ),
      stStationsParameter                   := ( rLaengeUebergroesseScheibe              := 4240,                            // Shuttle: ab dieser Scheibenlaenge gilt die Scheibe als uebergross [mm]
                                                 rMinGlasHoeheAutomatischenEintransport  := 500,                             // VSG: Mindesthoehe fuer automatischen Eintransport [mm]
                                                 rMinGlasLaengeAutomatischenEintransport := 500,                             // VSG: Mindestlaenge fuer automatischen Eintransport [mm]
                                                 wMaximaleAnzahlAktiverAuftraege := 1,                                       // derzeit ohne Funktion
                                                 rMinPosSwEsEingrenzung                  := 0.0,                             // Externer zusaetzlicher Software-Endschalter MIN; 0 = inaktiv; darf den MK-MIN nur weiter eingrenzen
                                                 rMaxPosSwEsEingrenzung                  := 0.0,                             // Externer zusaetzlicher Software-Endschalter MAX; 0 = inaktiv; darf den MK-MAX nur weiter eingrenzen
                                                 rPosFreigabePufferAusfahren             := 0.0                              // derzeit ohne Funktion
                                              ),
      // stFremdanlage
      stGlasdaten                           := [( rlMinGlasLaenge := 350,                                                    // minimal zulässige GlasLänge
                                                  rlMaxGlasLaenge := 2500,                                                   // maximale zulässige GlasLänge
                                                  rlMinGlasHoehe  := 190,                                                    // minimal zulässige GlasHöhe
                                                  rlMaxGlasHoehe  := 1800,                                                   // maximale zulässige GlasHöhe
                                                  rlMinGlasDicke  := 3,                                                    // minimal zulässige GlasDicke
                                                  rlMaxGlasDicke  := 12.76,                                                     // maximal zulaessige Glasdicke [mm]
                                                  rlLaengeMaxGlas := 0.0                                                     // maximal zulaessige Glaslaenge [mm]
                                               )]
      // astShuttleAnhaltenQuellen
    );

  apgMKStation203Glastransport : ARRAY[cWAND_1..cANZAHL_WAENDE] OF Parameter_Glastransport := [
    (
      rLaengeStation                        := 2600, // Länge der Station
      rScheibenabstand                      :=  300, // Der Abstand zwischen zwei Scheiben auf der Station
      rWegUeberEinlauf                      :=   50, // Weg ueber den Einlaufsensor hinaus [mm]
      rWegUeberAuslauf                      :=   50, // Weg ueber den Auslaufsensor hinaus [mm]
      rWegUeberSensorenSystemCheck          :=   15, // Der Weg der Ueber ein die Sensoren zum vermessen der Scheiben
      rUeberwachungAuslaufsensor            :=  500, // Ueberwachung des Auslaufsensors [Strecke in der der Auslaufsensor Frei / ueberfahren werden soll]
      rUeberwachungEinlaufsensor            :=  500, // Ueberwachung des Einlaufsensors [Strecke in der der Einlaufsensor Frei / ueberfahren werden soll]
      rWegUeberEinlaufEintransport          :=   30, // Eintransport vorwaerts: Abstand Scheibenhinterkante zum Einlaufsensor [mm]
      rWegUeberEinlaufAustransport          :=   50, // Lage Auf Einlauf: Scheibe liegt um diesen Weg auf dem Einlaufsensor [mm]
      rWegUeberAuslaufEintransport          :=   50, // Eintransport rueckwaerts: Abstand Scheibenhinterkante zum Auslaufsensor [mm]
      rWegUeberAuslaufAustransport          :=   50, // Lage Auf Auslauf: Weg ueber den Auslaufsensor hinaus [mm]
      rWegEinlaufsensorZuVorStopSensor      := 2400, // Beschreibt den Weg vum eine Scheibe beim EIntransport vom Einlaufsensor bis ueberden Vorabstopsensor zu verfahren
      rMesstoleranz                         :=   10, // Toleranz-Mass fuer die Scheibenlaengenmessung
      rMessstrecke                          := 2525, // Beschreibt die Strecke ziwischen 2 Sensoren die der Antrieb verfaehrt
      rWegstreckeBisZurVerzoegerung         := 1900  // Beschreibt die Strecke die gefahren werden soll bis der Antrieb abgebremst werden soll, dies gilt fuer Eintransportauftraege die das Bit "Letzte Scheibe" gesetzt haben
    )];

  apgMKStation203Kippen : ARRAY[cWAND_1..cANZAHL_WAENDE] OF Parameter_Kippen := [
    (
      tZeitlicheUeberwachungKippen          := TIME#5000MS, // [ms \ s] Verwendet fuer Antriebe die Ueber einen Schuetz angesteuert werden
      tZeitAntriebsfreigabeErhalten         := TIME#180S,   // [ms \ s] Energieeinsparrung: Zeiteinheit nach der die Antriebsfreigabe entzogen werden soll wenn keine Aktion ansteht [1 s = 1000 ms ]
      rToleranz                             := 0,           // Toleranz beim Entscheiden der aktuellen Position
      rPosition0Grad                        := 0,           // Waagerechte- Position 0 Grad: Position auf die die Station gehoben werden soll
      rPosition84Grad                       := 0,           // Senkrechte- Position 84 Grad: Position auf die die Station gehoben werden soll
      rPosition90Grad                       := 0,           // Senkrechte-Position 90 Grad : Position auf die die Station gesenkt werden soll
      rPosition96Grad                       := 0,           // Senkrechte-Position 96 Grad : Position auf die die Station gesenkt werden soll
      bKippenMitSchuetz                     := TRUE,        // Kippen per Umrichter oder Schütz
      rPosition88_5Grad                     := 0.0          // Senkrechte- Position 84 Grad: Position auf die die Station gehoben werden soll
    )];

   apgMKStation203Querfahrt : Parameter_Querfahrt :=
    (
      tZeitAntriebsfreigabeErhalten          := T#3M // Energieeinsparung: Zeit nach der die Antriebsfreigabe entzogen wird, wenn keine Aktion ansteht
    );

END_VAR
END_NAMESPACE

(* ---- Konfiguration_202.gvl ---- *)
(* METADATA
{
	"v3Meta": {
		"objectGuid": "5ca9fbcb-dcde-4398-ba5d-664b1abf1008"
	}
}
*)
{attribute 'allow_unqualified_access'}
NAMESPACE Konfiguration_202
VAR_CONFIG
//-------------------------------------------------------------------------------------------------
// KONFIGURATION: BAUSTEIN IO´s
//-------------------------------------------------------------------------------------------------
  // IO's GEBLAESE
  Globale_Bausteine.Foerderer202.Geblaese.in_bMotorschutzschalter_OK                 AT %MX1.1    : BOOL; // OPTION
  Globale_Bausteine.Foerderer202.Geblaese.out_bStarteGeblaese                        AT %MX2020.0 : BOOL; // OPTION

  // IO's KIPPEN
  Globale_Bausteine.Foerderer202.Kippen.in_bMotorstarter_OK                          AT %MX1.1    : BOOL; // OPTION
  Globale_Bausteine.Foerderer202.Kippen.in_bLS400V_OK                                AT %MX1.1    : BOOL; // OPTION
  Globale_Bausteine.Foerderer202.Kippen.in_bLSBremse_OK                              AT %MX1.1    : BOOL; // OPTION

  Globale_Bausteine.Foerderer202.Kippen.out_bKippen84Grad                            AT %MX2020.1 : BOOL; // OPTION
  Globale_Bausteine.Foerderer202.Kippen.out_bKippen90Grad                            AT %MX2020.2 : BOOL; // OPTION
  Globale_Bausteine.Foerderer202.Kippen.out_bBremseLoesen                            AT %MX2020.3 : BOOL; // OPTION
  Globale_Bausteine.Foerderer202.Kippen.out_bReset                                   AT %MX2020.4 : BOOL; // OPTION

  // IO's Hub
  Globale_Bausteine.Foerderer202.Hub.in_bLSBremse_OK                                 AT %MX1.1    : BOOL; // OPTION
  Globale_Bausteine.Foerderer202.Hub.in_bMotorstarter_OK                             AT %MX1.1    : BOOL; // OPTION
  Globale_Bausteine.Foerderer202.Hub.in_bLS400V_OK                                   AT %MX1.1    : BOOL; // OPTION
  Globale_Bausteine.Foerderer202.Hub.in_bSensorNichtOben                             AT %MX1.0    : BOOL; // OPTION
  Globale_Bausteine.Foerderer202.Hub.in_bSensorNichtUnten                            AT %MX1.1    : BOOL; // OPTION

  Globale_Bausteine.Foerderer202.Hub.out_bHubAbSetzen                                AT %MX2020.5 : BOOL; // OPTION
  Globale_Bausteine.Foerderer202.Hub.out_bHubAufSetzen                               AT %MX2020.6 : BOOL; // OPTION
  Globale_Bausteine.Foerderer202.Hub.out_bReset                                      AT %MX2020.7 : BOOL; // OPTION
  Globale_Bausteine.Foerderer202.Hub.out_bBremseLoesen                               AT %MX2021.0 : BOOL; // OPTION

  // IO's RÖLLCHENLEISTE
  Globale_Bausteine.Foerderer202.Roellchenleiste.in_bStatusZylinder1Ausgefahren      AT %MX1.0    : BOOL; // OPTION
  Globale_Bausteine.Foerderer202.Roellchenleiste.in_bStatusZylinder1Eingefahren      AT %MX1.0    : BOOL; // OPTION
  Globale_Bausteine.Foerderer202.Roellchenleiste.in_bStatusZylinder2Ausgefahren      AT %MX1.0    : BOOL; // OPTION
  Globale_Bausteine.Foerderer202.Roellchenleiste.in_bStatusZylinder2Eingefahren      AT %MX1.0    : BOOL; // OPTION

  Globale_Bausteine.Foerderer202.Roellchenleiste.out_bZylinder1Ausfahren             AT %MX2021.1 : BOOL; // OPTION
  Globale_Bausteine.Foerderer202.Roellchenleiste.out_bZylinder1Einfahren             AT %MX2021.2 : BOOL; // OPTION
  Globale_Bausteine.Foerderer202.Roellchenleiste.out_bZylinder2Ausfahren             AT %MX2021.3 : BOOL; // OPTION
  Globale_Bausteine.Foerderer202.Roellchenleiste.out_bZylinder2Einfahren             AT %MX2021.4 : BOOL; // OPTION

  // IO's WANDVERSTELLUNG
  Globale_Bausteine.Foerderer202.Wandverstellung.in_bStatusZylinder1Ausgefahren      AT %MX1.0    : BOOL; // OPTION
  Globale_Bausteine.Foerderer202.Wandverstellung.in_bStatusZylinder1Eingefahren      AT %MX1.0    : BOOL; // OPTION
  Globale_Bausteine.Foerderer202.Wandverstellung.in_bStatusZylinder2Ausgefahren      AT %MX1.0    : BOOL; // OPTION
  Globale_Bausteine.Foerderer202.Wandverstellung.in_bStatusZylinder2Eingefahren      AT %MX1.0    : BOOL; // OPTION

  Globale_Bausteine.Foerderer202.Wandverstellung.out_bZylinder1Ausfahren             AT %MX2021.5 : BOOL; // OPTION
  Globale_Bausteine.Foerderer202.Wandverstellung.out_bZylinder1Einfahren             AT %MX2021.6 : BOOL; // OPTION
  Globale_Bausteine.Foerderer202.Wandverstellung.out_bZylinder2Ausfahren             AT %MX2021.7 : BOOL; // OPTION
  Globale_Bausteine.Foerderer202.Wandverstellung.out_bZylinder2Einfahren             AT %MX2022.0 : BOOL; // OPTION

END_VAR

END_NAMESPACE

(* ---- Konfiguration_203.gvl ---- *)
(* METADATA
{
	"v3Meta": {
		"objectGuid": "2bacb3a2-0057-4448-8d3c-3d597e0de1a8"
	}
}
*)
{attribute 'allow_unqualified_access'}
NAMESPACE Konfiguration_203
VAR_CONFIG
//-------------------------------------------------------------------------------------------------
// KONFIGURATION: BAUSTEIN IO´s
//-------------------------------------------------------------------------------------------------
  // IO's GEBLAESE
  Globale_Bausteine.Foerderer203.Geblaese.in_bMotorschutzschalter_OK                 AT %MX1.1    : BOOL; // OPTION
  Globale_Bausteine.Foerderer203.Geblaese.out_bStarteGeblaese                        AT %MX2030.0 : BOOL; // OPTION

  // IO's KIPPEN
  Globale_Bausteine.Foerderer203.Kippen.in_bMotorstarter_OK                          AT %MX1.1    : BOOL; // OPTION
  Globale_Bausteine.Foerderer203.Kippen.in_bLS400V_OK                                AT %MX1.1    : BOOL; // OPTION
  Globale_Bausteine.Foerderer203.Kippen.in_bLSBremse_OK                              AT %MX1.1    : BOOL; // OPTION

  Globale_Bausteine.Foerderer203.Kippen.out_bKippen84Grad                            AT %MX2030.1 : BOOL; // OPTION
  Globale_Bausteine.Foerderer203.Kippen.out_bKippen90Grad                            AT %MX2030.2 : BOOL; // OPTION
  Globale_Bausteine.Foerderer203.Kippen.out_bBremseLoesen                            AT %MX2030.3 : BOOL; // OPTION
  Globale_Bausteine.Foerderer203.Kippen.out_bReset                                   AT %MX2030.4 : BOOL; // OPTION

  // IO's Hub
  Globale_Bausteine.Foerderer203.Hub.in_bLSBremse_OK                                 AT %MX1.1    : BOOL; // OPTION
  Globale_Bausteine.Foerderer203.Hub.in_bMotorstarter_OK                             AT %MX1.1    : BOOL; // OPTION
  Globale_Bausteine.Foerderer203.Hub.in_bLS400V_OK                                   AT %MX1.1    : BOOL; // OPTION
  Globale_Bausteine.Foerderer203.Hub.in_bSensorNichtOben                             AT %MX1.0    : BOOL; // OPTION
  Globale_Bausteine.Foerderer203.Hub.in_bSensorNichtUnten                            AT %MX1.1    : BOOL; // OPTION

  Globale_Bausteine.Foerderer203.Hub.out_bHubAbSetzen                                AT %MX2030.5 : BOOL; // OPTION
  Globale_Bausteine.Foerderer203.Hub.out_bHubAufSetzen                               AT %MX2030.6 : BOOL; // OPTION
  Globale_Bausteine.Foerderer203.Hub.out_bReset                                      AT %MX2030.7 : BOOL; // OPTION
  Globale_Bausteine.Foerderer203.Hub.out_bBremseLoesen                               AT %MX2031.0 : BOOL; // OPTION

  // IO's RÖLLCHENLEISTE
  Globale_Bausteine.Foerderer203.Roellchenleiste.in_bStatusZylinder1Ausgefahren      AT %MX1.0    : BOOL; // OPTION
  Globale_Bausteine.Foerderer203.Roellchenleiste.in_bStatusZylinder1Eingefahren      AT %MX1.0    : BOOL; // OPTION
  Globale_Bausteine.Foerderer203.Roellchenleiste.in_bStatusZylinder2Ausgefahren      AT %MX1.0    : BOOL; // OPTION
  Globale_Bausteine.Foerderer203.Roellchenleiste.in_bStatusZylinder2Eingefahren      AT %MX1.0    : BOOL; // OPTION

  Globale_Bausteine.Foerderer203.Roellchenleiste.out_bZylinder1Ausfahren             AT %MX2031.1 : BOOL; // OPTION
  Globale_Bausteine.Foerderer203.Roellchenleiste.out_bZylinder1Einfahren             AT %MX2031.2 : BOOL; // OPTION
  Globale_Bausteine.Foerderer203.Roellchenleiste.out_bZylinder2Ausfahren             AT %MX2031.3 : BOOL; // OPTION
  Globale_Bausteine.Foerderer203.Roellchenleiste.out_bZylinder2Einfahren             AT %MX2031.4 : BOOL; // OPTION

  // IO's WANDVERSTELLUNG
  Globale_Bausteine.Foerderer203.Wandverstellung.in_bStatusZylinder1Ausgefahren      AT %MX1.0    : BOOL; // OPTION
  Globale_Bausteine.Foerderer203.Wandverstellung.in_bStatusZylinder1Eingefahren      AT %MX1.0    : BOOL; // OPTION
  Globale_Bausteine.Foerderer203.Wandverstellung.in_bStatusZylinder2Ausgefahren      AT %MX1.0    : BOOL; // OPTION
  Globale_Bausteine.Foerderer203.Wandverstellung.in_bStatusZylinder2Eingefahren      AT %MX1.0    : BOOL; // OPTION

  Globale_Bausteine.Foerderer203.Wandverstellung.out_bZylinder1Ausfahren             AT %MX2031.5 : BOOL; // OPTION
  Globale_Bausteine.Foerderer203.Wandverstellung.out_bZylinder1Einfahren             AT %MX2031.6 : BOOL; // OPTION
  Globale_Bausteine.Foerderer203.Wandverstellung.out_bZylinder2Ausfahren             AT %MX2031.7 : BOOL; // OPTION
  Globale_Bausteine.Foerderer203.Wandverstellung.out_bZylinder2Einfahren             AT %MX2032.0 : BOOL; // OPTION

END_VAR

END_NAMESPACE
